(* IEC 61131-3 sources: s7-to-codesys/tests/POUs/Scenarios/FB_Motor_ScenarioTest, 8 files *)

(* ---- FB_Motor_ScenarioTest.decl.st ---- *)
// AUTO-GENERATED — не редактировать: s7conv gen-tests, сценарии scenarios/FB_Motor.csv
// Правка — в CSV (scenarios/README.md), затем python -m s7conv build-corpus.
// Назначение: тесты поведения сконвертированного FB_Motor по сценариям CSV (сценариев: 7, строк: 52):
//             один метод-тест на сценарий, строки — по порядку с моделируемым временем GVL_S7Clock.
//             Ожидаемые значения — из CSV (эталонные модели по описанию логики блока), не из
//             результата конвертации.
// Автор:      s7conv 0.1.0 (сгенерировано)
// Версия:     не указана
// Документ:   scenarios/README.md, docs/methodology.md, раздел «Проверка поведения»
FUNCTION_BLOCK FB_Motor_ScenarioTest EXTENDS coUnit.FB_TestSuite
VAR
    fbAutoStartOk : FB_Motor;  // свой экземпляр на сценарий
    xAutoStartOkDone : BOOL;  // сценарий выполнен (выполняется один раз)
    fbNoFeedbackTimeout : FB_Motor;  // свой экземпляр на сценарий
    xNoFeedbackTimeoutDone : BOOL;  // сценарий выполнен (выполняется один раз)
    fbFeedbackLost : FB_Motor;  // свой экземпляр на сценарий
    xFeedbackLostDone : BOOL;  // сценарий выполнен (выполняется один раз)
    fbUnexpectedFeedback : FB_Motor;  // свой экземпляр на сценарий
    xUnexpectedFeedbackDone : BOOL;  // сценарий выполнен (выполняется один раз)
    fbThermalTripManual : FB_Motor;  // свой экземпляр на сценарий
    xThermalTripManualDone : BOOL;  // сценарий выполнен (выполняется один раз)
    fbBumplessAutoToManual : FB_Motor;  // свой экземпляр на сценарий
    xBumplessAutoToManualDone : BOOL;  // сценарий выполнен (выполняется один раз)
    fbCustomFeedbackTime : FB_Motor;  // свой экземпляр на сценарий
    xCustomFeedbackTimeDone : BOOL;  // сценарий выполнен (выполняется один раз)
END_VAR

(* ---- AutoStartOk.method.impl.st ---- *)
// AUTO-GENERATED — не редактировать: scenarios/FB_Motor.csv, сценарий AutoStartOk
coUnit.TEST('AutoStartOk');
IF NOT xAutoStartOkDone THEN
    xAutoStartOkDone := TRUE;
    GVL_S7Clock.xSimulation := TRUE;

    // #1, t = 0 мс — авто, команды нет
    GVL_S7Clock.tSimNow := T#0MS;
    fbAutoStartOk.autoMode := TRUE;
    fbAutoStartOk.autoStart := FALSE;
    fbAutoStartOk.manStart := FALSE;
    fbAutoStartOk.manStop := FALSE;
    fbAutoStartOk.feedback := FALSE;
    fbAutoStartOk.thermalOk := TRUE;
    fbAutoStartOk.reset := FALSE;
    fbAutoStartOk.feedbackTime := T#3000MS;
    fbAutoStartOk();
    AssertEquals_BOOL(Expected := FALSE, Actual := fbAutoStartOk.runCmd, Message := 'AutoStartOk#1 runCmd');
    AssertEquals_BOOL(Expected := FALSE, Actual := fbAutoStartOk.fault, Message := 'AutoStartOk#1 fault');
    AssertEquals_BOOL(Expected := FALSE,
                      Actual := fbAutoStartOk.status.running,
                      Message := 'AutoStartOk#1 status.running');
    AssertEquals_BOOL(Expected := FALSE, Actual := fbAutoStartOk.status.fault, Message := 'AutoStartOk#1 status.fault');
    AssertEquals_BOOL(Expected := TRUE,
                      Actual := fbAutoStartOk.status.autoMode,
                      Message := 'AutoStartOk#1 status.autoMode');
    AssertEquals_INT(Expected := 0,
                     Actual := fbAutoStartOk.status.faultCode,
                     Message := 'AutoStartOk#1 status.faultCode');
    AssertEquals_DINT(Expected := 0,
                      Actual := fbAutoStartOk.status.startCount,
                      Message := 'AutoStartOk#1 status.startCount');

    // #2, t = 100 мс — пуск: runCmd, пуск №1; таймер рассогласования запущен
    GVL_S7Clock.tSimNow := T#100MS;
    fbAutoStartOk.autoStart := TRUE;
    fbAutoStartOk();
    AssertEquals_BOOL(Expected := TRUE, Actual := fbAutoStartOk.runCmd, Message := 'AutoStartOk#2 runCmd');
    AssertEquals_BOOL(Expected := FALSE, Actual := fbAutoStartOk.fault, Message := 'AutoStartOk#2 fault');
    AssertEquals_BOOL(Expected := FALSE,
                      Actual := fbAutoStartOk.status.running,
                      Message := 'AutoStartOk#2 status.running');
    AssertEquals_BOOL(Expected := FALSE, Actual := fbAutoStartOk.status.fault, Message := 'AutoStartOk#2 status.fault');
    AssertEquals_BOOL(Expected := TRUE,
                      Actual := fbAutoStartOk.status.autoMode,
                      Message := 'AutoStartOk#2 status.autoMode');
    AssertEquals_INT(Expected := 0,
                     Actual := fbAutoStartOk.status.faultCode,
                     Message := 'AutoStartOk#2 status.faultCode');
    AssertEquals_DINT(Expected := 1,
                      Actual := fbAutoStartOk.status.startCount,
                      Message := 'AutoStartOk#2 status.startCount');

    // #3, t = 1100 мс — обратная связь через 1 с: работает
    GVL_S7Clock.tSimNow := T#1100MS;
    fbAutoStartOk.feedback := TRUE;
    fbAutoStartOk();
    AssertEquals_BOOL(Expected := TRUE, Actual := fbAutoStartOk.runCmd, Message := 'AutoStartOk#3 runCmd');
    AssertEquals_BOOL(Expected := FALSE, Actual := fbAutoStartOk.fault, Message := 'AutoStartOk#3 fault');
    AssertEquals_BOOL(Expected := TRUE,
                      Actual := fbAutoStartOk.status.running,
                      Message := 'AutoStartOk#3 status.running');
    AssertEquals_BOOL(Expected := FALSE, Actual := fbAutoStartOk.status.fault, Message := 'AutoStartOk#3 status.fault');
    AssertEquals_BOOL(Expected := TRUE,
                      Actual := fbAutoStartOk.status.autoMode,
                      Message := 'AutoStartOk#3 status.autoMode');
    AssertEquals_INT(Expected := 0,
                     Actual := fbAutoStartOk.status.faultCode,
                     Message := 'AutoStartOk#3 status.faultCode');
    AssertEquals_DINT(Expected := 1,
                      Actual := fbAutoStartOk.status.startCount,
                      Message := 'AutoStartOk#3 status.startCount');

    // #4, t = 5000 мс — работает, аварии нет
    GVL_S7Clock.tSimNow := T#5000MS;
    fbAutoStartOk();
    AssertEquals_BOOL(Expected := TRUE, Actual := fbAutoStartOk.runCmd, Message := 'AutoStartOk#4 runCmd');
    AssertEquals_BOOL(Expected := FALSE, Actual := fbAutoStartOk.fault, Message := 'AutoStartOk#4 fault');
    AssertEquals_BOOL(Expected := TRUE,
                      Actual := fbAutoStartOk.status.running,
                      Message := 'AutoStartOk#4 status.running');
    AssertEquals_BOOL(Expected := FALSE, Actual := fbAutoStartOk.status.fault, Message := 'AutoStartOk#4 status.fault');
    AssertEquals_BOOL(Expected := TRUE,
                      Actual := fbAutoStartOk.status.autoMode,
                      Message := 'AutoStartOk#4 status.autoMode');
    AssertEquals_INT(Expected := 0,
                     Actual := fbAutoStartOk.status.faultCode,
                     Message := 'AutoStartOk#4 status.faultCode');
    AssertEquals_DINT(Expected := 1,
                      Actual := fbAutoStartOk.status.startCount,
                      Message := 'AutoStartOk#4 status.startCount');

    // #5, t = 5100 мс — стоп: runCmd снят, контактор ещё держит — рассогласование
    GVL_S7Clock.tSimNow := T#5100MS;
    fbAutoStartOk.autoStart := FALSE;
    fbAutoStartOk();
    AssertEquals_BOOL(Expected := FALSE, Actual := fbAutoStartOk.runCmd, Message := 'AutoStartOk#5 runCmd');
    AssertEquals_BOOL(Expected := FALSE, Actual := fbAutoStartOk.fault, Message := 'AutoStartOk#5 fault');
    AssertEquals_BOOL(Expected := FALSE,
                      Actual := fbAutoStartOk.status.running,
                      Message := 'AutoStartOk#5 status.running');
    AssertEquals_BOOL(Expected := FALSE, Actual := fbAutoStartOk.status.fault, Message := 'AutoStartOk#5 status.fault');
    AssertEquals_BOOL(Expected := TRUE,
                      Actual := fbAutoStartOk.status.autoMode,
                      Message := 'AutoStartOk#5 status.autoMode');
    AssertEquals_INT(Expected := 0,
                     Actual := fbAutoStartOk.status.faultCode,
                     Message := 'AutoStartOk#5 status.faultCode');
    AssertEquals_DINT(Expected := 1,
                      Actual := fbAutoStartOk.status.startCount,
                      Message := 'AutoStartOk#5 status.startCount');

    // #6, t = 6000 мс — обратная связь пропала через 0.9 с — нормальный останов
    GVL_S7Clock.tSimNow := T#6000MS;
    fbAutoStartOk.feedback := FALSE;
    fbAutoStartOk();
    AssertEquals_BOOL(Expected := FALSE, Actual := fbAutoStartOk.runCmd, Message := 'AutoStartOk#6 runCmd');
    AssertEquals_BOOL(Expected := FALSE, Actual := fbAutoStartOk.fault, Message := 'AutoStartOk#6 fault');
    AssertEquals_BOOL(Expected := FALSE,
                      Actual := fbAutoStartOk.status.running,
                      Message := 'AutoStartOk#6 status.running');
    AssertEquals_BOOL(Expected := FALSE, Actual := fbAutoStartOk.status.fault, Message := 'AutoStartOk#6 status.fault');
    AssertEquals_BOOL(Expected := TRUE,
                      Actual := fbAutoStartOk.status.autoMode,
                      Message := 'AutoStartOk#6 status.autoMode');
    AssertEquals_INT(Expected := 0,
                     Actual := fbAutoStartOk.status.faultCode,
                     Message := 'AutoStartOk#6 status.faultCode');
    AssertEquals_DINT(Expected := 1,
                      Actual := fbAutoStartOk.status.startCount,
                      Message := 'AutoStartOk#6 status.startCount');

    // #7, t = 9500 мс — покой
    GVL_S7Clock.tSimNow := T#9500MS;
    fbAutoStartOk();
    AssertEquals_BOOL(Expected := FALSE, Actual := fbAutoStartOk.runCmd, Message := 'AutoStartOk#7 runCmd');
    AssertEquals_BOOL(Expected := FALSE, Actual := fbAutoStartOk.fault, Message := 'AutoStartOk#7 fault');
    AssertEquals_BOOL(Expected := FALSE,
                      Actual := fbAutoStartOk.status.running,
                      Message := 'AutoStartOk#7 status.running');
    AssertEquals_BOOL(Expected := FALSE, Actual := fbAutoStartOk.status.fault, Message := 'AutoStartOk#7 status.fault');
    AssertEquals_BOOL(Expected := TRUE,
                      Actual := fbAutoStartOk.status.autoMode,
                      Message := 'AutoStartOk#7 status.autoMode');
    AssertEquals_INT(Expected := 0,
                     Actual := fbAutoStartOk.status.faultCode,
                     Message := 'AutoStartOk#7 status.faultCode');
    AssertEquals_DINT(Expected := 1,
                      Actual := fbAutoStartOk.status.startCount,
                      Message := 'AutoStartOk#7 status.startCount');

    GVL_S7Clock.xSimulation := FALSE;
END_IF
coUnit.TEST_FINISHED();

(* ---- BumplessAutoToManual.method.impl.st ---- *)
// AUTO-GENERATED — не редактировать: scenarios/FB_Motor.csv, сценарий BumplessAutoToManual
coUnit.TEST('BumplessAutoToManual');
IF NOT xBumplessAutoToManualDone THEN
    xBumplessAutoToManualDone := TRUE;
    GVL_S7Clock.xSimulation := TRUE;

    // #1, t = 0 мс — авто, пуск №1
    GVL_S7Clock.tSimNow := T#0MS;
    fbBumplessAutoToManual.autoMode := TRUE;
    fbBumplessAutoToManual.autoStart := TRUE;
    fbBumplessAutoToManual.manStart := FALSE;
    fbBumplessAutoToManual.manStop := FALSE;
    fbBumplessAutoToManual.feedback := FALSE;
    fbBumplessAutoToManual.thermalOk := TRUE;
    fbBumplessAutoToManual.reset := FALSE;
    fbBumplessAutoToManual.feedbackTime := T#3000MS;
    fbBumplessAutoToManual();
    AssertEquals_BOOL(Expected := TRUE,
                      Actual := fbBumplessAutoToManual.runCmd,
                      Message := 'BumplessAutoToManual#1 runCmd');
    AssertEquals_BOOL(Expected := FALSE,
                      Actual := fbBumplessAutoToManual.fault,
                      Message := 'BumplessAutoToManual#1 fault');
    AssertEquals_BOOL(Expected := FALSE,
                      Actual := fbBumplessAutoToManual.status.running,
                      Message := 'BumplessAutoToManual#1 status.running');
    AssertEquals_BOOL(Expected := FALSE,
                      Actual := fbBumplessAutoToManual.status.fault,
                      Message := 'BumplessAutoToManual#1 status.fault');
    AssertEquals_BOOL(Expected := TRUE,
                      Actual := fbBumplessAutoToManual.status.autoMode,
                      Message := 'BumplessAutoToManual#1 status.autoMode');
    AssertEquals_INT(Expected := 0,
                     Actual := fbBumplessAutoToManual.status.faultCode,
                     Message := 'BumplessAutoToManual#1 status.faultCode');
    AssertEquals_DINT(Expected := 1,
                      Actual := fbBumplessAutoToManual.status.startCount,
                      Message := 'BumplessAutoToManual#1 status.startCount');

    // #2, t = 500 мс — работает
    GVL_S7Clock.tSimNow := T#500MS;
    fbBumplessAutoToManual.feedback := TRUE;
    fbBumplessAutoToManual();
    AssertEquals_BOOL(Expected := TRUE,
                      Actual := fbBumplessAutoToManual.runCmd,
                      Message := 'BumplessAutoToManual#2 runCmd');
    AssertEquals_BOOL(Expected := FALSE,
                      Actual := fbBumplessAutoToManual.fault,
                      Message := 'BumplessAutoToManual#2 fault');
    AssertEquals_BOOL(Expected := TRUE,
                      Actual := fbBumplessAutoToManual.status.running,
                      Message := 'BumplessAutoToManual#2 status.running');
    AssertEquals_BOOL(Expected := FALSE,
                      Actual := fbBumplessAutoToManual.status.fault,
                      Message := 'BumplessAutoToManual#2 status.fault');
    AssertEquals_BOOL(Expected := TRUE,
                      Actual := fbBumplessAutoToManual.status.autoMode,
                      Message := 'BumplessAutoToManual#2 status.autoMode');
    AssertEquals_INT(Expected := 0,
                     Actual := fbBumplessAutoToManual.status.faultCode,
                     Message := 'BumplessAutoToManual#2 status.faultCode');
    AssertEquals_DINT(Expected := 1,
                      Actual := fbBumplessAutoToManual.status.startCount,
                      Message := 'BumplessAutoToManual#2 status.startCount');

    // #3, t = 1000 мс — в ручной: защёлка следила за авто — продолжает работать
    GVL_S7Clock.tSimNow := T#1000MS;
    fbBumplessAutoToManual.autoMode := FALSE;
    fbBumplessAutoToManual();
    AssertEquals_BOOL(Expected := TRUE,
                      Actual := fbBumplessAutoToManual.runCmd,
                      Message := 'BumplessAutoToManual#3 runCmd');
    AssertEquals_BOOL(Expected := FALSE,
                      Actual := fbBumplessAutoToManual.fault,
                      Message := 'BumplessAutoToManual#3 fault');
    AssertEquals_BOOL(Expected := TRUE,
                      Actual := fbBumplessAutoToManual.status.running,
                      Message := 'BumplessAutoToManual#3 status.running');
    AssertEquals_BOOL(Expected := FALSE,
                      Actual := fbBumplessAutoToManual.status.fault,
                      Message := 'BumplessAutoToManual#3 status.fault');
    AssertEquals_BOOL(Expected := FALSE,
                      Actual := fbBumplessAutoToManual.status.autoMode,
                      Message := 'BumplessAutoToManual#3 status.autoMode');
    AssertEquals_INT(Expected := 0,
                     Actual := fbBumplessAutoToManual.status.faultCode,
                     Message := 'BumplessAutoToManual#3 status.faultCode');
    AssertEquals_DINT(Expected := 1,
                      Actual := fbBumplessAutoToManual.status.startCount,
                      Message := 'BumplessAutoToManual#3 status.startCount');

    // #4, t = 2000 мс — стоп оператором
    GVL_S7Clock.tSimNow := T#2000MS;
    fbBumplessAutoToManual.manStop := TRUE;
    fbBumplessAutoToManual();
    AssertEquals_BOOL(Expected := FALSE,
                      Actual := fbBumplessAutoToManual.runCmd,
                      Message := 'BumplessAutoToManual#4 runCmd');
    AssertEquals_BOOL(Expected := FALSE,
                      Actual := fbBumplessAutoToManual.fault,
                      Message := 'BumplessAutoToManual#4 fault');
    AssertEquals_BOOL(Expected := FALSE,
                      Actual := fbBumplessAutoToManual.status.running,
                      Message := 'BumplessAutoToManual#4 status.running');
    AssertEquals_BOOL(Expected := FALSE,
                      Actual := fbBumplessAutoToManual.status.fault,
                      Message := 'BumplessAutoToManual#4 status.fault');
    AssertEquals_BOOL(Expected := FALSE,
                      Actual := fbBumplessAutoToManual.status.autoMode,
                      Message := 'BumplessAutoToManual#4 status.autoMode');
    AssertEquals_INT(Expected := 0,
                     Actual := fbBumplessAutoToManual.status.faultCode,
                     Message := 'BumplessAutoToManual#4 status.faultCode');
    AssertEquals_DINT(Expected := 1,
                      Actual := fbBumplessAutoToManual.status.startCount,
                      Message := 'BumplessAutoToManual#4 status.startCount');

    // #5, t = 2500 мс — остановлен
    GVL_S7Clock.tSimNow := T#2500MS;
    fbBumplessAutoToManual.manStop := FALSE;
    fbBumplessAutoToManual.feedback := FALSE;
    fbBumplessAutoToManual();
    AssertEquals_BOOL(Expected := FALSE,
                      Actual := fbBumplessAutoToManual.runCmd,
                      Message := 'BumplessAutoToManual#5 runCmd');
    AssertEquals_BOOL(Expected := FALSE,
                      Actual := fbBumplessAutoToManual.fault,
                      Message := 'BumplessAutoToManual#5 fault');
    AssertEquals_BOOL(Expected := FALSE,
                      Actual := fbBumplessAutoToManual.status.running,
                      Message := 'BumplessAutoToManual#5 status.running');
    AssertEquals_BOOL(Expected := FALSE,
                      Actual := fbBumplessAutoToManual.status.fault,
                      Message := 'BumplessAutoToManual#5 status.fault');
    AssertEquals_BOOL(Expected := FALSE,
                      Actual := fbBumplessAutoToManual.status.autoMode,
                      Message := 'BumplessAutoToManual#5 status.autoMode');
    AssertEquals_INT(Expected := 0,
                     Actual := fbBumplessAutoToManual.status.faultCode,
                     Message := 'BumplessAutoToManual#5 status.faultCode');
    AssertEquals_DINT(Expected := 1,
                      Actual := fbBumplessAutoToManual.status.startCount,
                      Message := 'BumplessAutoToManual#5 status.startCount');

    // #6, t = 3000 мс — в авто без запроса
    GVL_S7Clock.tSimNow := T#3000MS;
    fbBumplessAutoToManual.autoMode := TRUE;
    fbBumplessAutoToManual.autoStart := FALSE;
    fbBumplessAutoToManual();
    AssertEquals_BOOL(Expected := FALSE,
                      Actual := fbBumplessAutoToManual.runCmd,
                      Message := 'BumplessAutoToManual#6 runCmd');
    AssertEquals_BOOL(Expected := FALSE,
                      Actual := fbBumplessAutoToManual.fault,
                      Message := 'BumplessAutoToManual#6 fault');
    AssertEquals_BOOL(Expected := FALSE,
                      Actual := fbBumplessAutoToManual.status.running,
                      Message := 'BumplessAutoToManual#6 status.running');
    AssertEquals_BOOL(Expected := FALSE,
                      Actual := fbBumplessAutoToManual.status.fault,
                      Message := 'BumplessAutoToManual#6 status.fault');
    AssertEquals_BOOL(Expected := TRUE,
                      Actual := fbBumplessAutoToManual.status.autoMode,
                      Message := 'BumplessAutoToManual#6 status.autoMode');
    AssertEquals_INT(Expected := 0,
                     Actual := fbBumplessAutoToManual.status.faultCode,
                     Message := 'BumplessAutoToManual#6 status.faultCode');
    AssertEquals_DINT(Expected := 1,
                      Actual := fbBumplessAutoToManual.status.startCount,
                      Message := 'BumplessAutoToManual#6 status.startCount');

    // #7, t = 3500 мс — запрос авто: пуск №2
    GVL_S7Clock.tSimNow := T#3500MS;
    fbBumplessAutoToManual.autoStart := TRUE;
    fbBumplessAutoToManual();
    AssertEquals_BOOL(Expected := TRUE,
                      Actual := fbBumplessAutoToManual.runCmd,
                      Message := 'BumplessAutoToManual#7 runCmd');
    AssertEquals_BOOL(Expected := FALSE,
                      Actual := fbBumplessAutoToManual.fault,
                      Message := 'BumplessAutoToManual#7 fault');
    AssertEquals_BOOL(Expected := FALSE,
                      Actual := fbBumplessAutoToManual.status.running,
                      Message := 'BumplessAutoToManual#7 status.running');
    AssertEquals_BOOL(Expected := FALSE,
                      Actual := fbBumplessAutoToManual.status.fault,
                      Message := 'BumplessAutoToManual#7 status.fault');
    AssertEquals_BOOL(Expected := TRUE,
                      Actual := fbBumplessAutoToManual.status.autoMode,
                      Message := 'BumplessAutoToManual#7 status.autoMode');
    AssertEquals_INT(Expected := 0,
                     Actual := fbBumplessAutoToManual.status.faultCode,
                     Message := 'BumplessAutoToManual#7 status.faultCode');
    AssertEquals_DINT(Expected := 2,
                      Actual := fbBumplessAutoToManual.status.startCount,
                      Message := 'BumplessAutoToManual#7 status.startCount');

    // #8, t = 4000 мс — работает
    GVL_S7Clock.tSimNow := T#4000MS;
    fbBumplessAutoToManual.feedback := TRUE;
    fbBumplessAutoToManual();
    AssertEquals_BOOL(Expected := TRUE,
                      Actual := fbBumplessAutoToManual.runCmd,
                      Message := 'BumplessAutoToManual#8 runCmd');
    AssertEquals_BOOL(Expected := FALSE,
                      Actual := fbBumplessAutoToManual.fault,
                      Message := 'BumplessAutoToManual#8 fault');
    AssertEquals_BOOL(Expected := TRUE,
                      Actual := fbBumplessAutoToManual.status.running,
                      Message := 'BumplessAutoToManual#8 status.running');
    AssertEquals_BOOL(Expected := FALSE,
                      Actual := fbBumplessAutoToManual.status.fault,
                      Message := 'BumplessAutoToManual#8 status.fault');
    AssertEquals_BOOL(Expected := TRUE,
                      Actual := fbBumplessAutoToManual.status.autoMode,
                      Message := 'BumplessAutoToManual#8 status.autoMode');
    AssertEquals_INT(Expected := 0,
                     Actual := fbBumplessAutoToManual.status.faultCode,
                     Message := 'BumplessAutoToManual#8 status.faultCode');
    AssertEquals_DINT(Expected := 2,
                      Actual := fbBumplessAutoToManual.status.startCount,
                      Message := 'BumplessAutoToManual#8 status.startCount');

    GVL_S7Clock.xSimulation := FALSE;
END_IF
coUnit.TEST_FINISHED();

(* ---- CustomFeedbackTime.method.impl.st ---- *)
// AUTO-GENERATED — не редактировать: scenarios/FB_Motor.csv, сценарий CustomFeedbackTime
coUnit.TEST('CustomFeedbackTime');
IF NOT xCustomFeedbackTimeDone THEN
    xCustomFeedbackTimeDone := TRUE;
    GVL_S7Clock.xSimulation := TRUE;

    // #1, t = 0 мс — пуск, feedbackTime 5 с
    GVL_S7Clock.tSimNow := T#0MS;
    fbCustomFeedbackTime.autoMode := TRUE;
    fbCustomFeedbackTime.autoStart := TRUE;
    fbCustomFeedbackTime.manStart := FALSE;
    fbCustomFeedbackTime.manStop := FALSE;
    fbCustomFeedbackTime.feedback := FALSE;
    fbCustomFeedbackTime.thermalOk := TRUE;
    fbCustomFeedbackTime.reset := FALSE;
    fbCustomFeedbackTime.feedbackTime := T#5000MS;
    fbCustomFeedbackTime();
    AssertEquals_BOOL(Expected := TRUE,
                      Actual := fbCustomFeedbackTime.runCmd,
                      Message := 'CustomFeedbackTime#1 runCmd');
    AssertEquals_BOOL(Expected := FALSE, Actual := fbCustomFeedbackTime.fault, Message := 'CustomFeedbackTime#1 fault');
    AssertEquals_BOOL(Expected := FALSE,
                      Actual := fbCustomFeedbackTime.status.running,
                      Message := 'CustomFeedbackTime#1 status.running');
    AssertEquals_BOOL(Expected := FALSE,
                      Actual := fbCustomFeedbackTime.status.fault,
                      Message := 'CustomFeedbackTime#1 status.fault');
    AssertEquals_BOOL(Expected := TRUE,
                      Actual := fbCustomFeedbackTime.status.autoMode,
                      Message := 'CustomFeedbackTime#1 status.autoMode');
    AssertEquals_INT(Expected := 0,
                     Actual := fbCustomFeedbackTime.status.faultCode,
                     Message := 'CustomFeedbackTime#1 status.faultCode');
    AssertEquals_DINT(Expected := 1,
                      Actual := fbCustomFeedbackTime.status.startCount,
                      Message := 'CustomFeedbackTime#1 status.startCount');

    // #2, t = 4500 мс — обратная связь через 4.5 с — аварии нет
    GVL_S7Clock.tSimNow := T#4500MS;
    fbCustomFeedbackTime.feedback := TRUE;
    fbCustomFeedbackTime();
    AssertEquals_BOOL(Expected := TRUE,
                      Actual := fbCustomFeedbackTime.runCmd,
                      Message := 'CustomFeedbackTime#2 runCmd');
    AssertEquals_BOOL(Expected := FALSE, Actual := fbCustomFeedbackTime.fault, Message := 'CustomFeedbackTime#2 fault');
    AssertEquals_BOOL(Expected := TRUE,
                      Actual := fbCustomFeedbackTime.status.running,
                      Message := 'CustomFeedbackTime#2 status.running');
    AssertEquals_BOOL(Expected := FALSE,
                      Actual := fbCustomFeedbackTime.status.fault,
                      Message := 'CustomFeedbackTime#2 status.fault');
    AssertEquals_BOOL(Expected := TRUE,
                      Actual := fbCustomFeedbackTime.status.autoMode,
                      Message := 'CustomFeedbackTime#2 status.autoMode');
    AssertEquals_INT(Expected := 0,
                     Actual := fbCustomFeedbackTime.status.faultCode,
                     Message := 'CustomFeedbackTime#2 status.faultCode');
    AssertEquals_DINT(Expected := 1,
                      Actual := fbCustomFeedbackTime.status.startCount,
                      Message := 'CustomFeedbackTime#2 status.startCount');

    // #3, t = 6000 мс — работает
    GVL_S7Clock.tSimNow := T#6000MS;
    fbCustomFeedbackTime();
    AssertEquals_BOOL(Expected := TRUE,
                      Actual := fbCustomFeedbackTime.runCmd,
                      Message := 'CustomFeedbackTime#3 runCmd');
    AssertEquals_BOOL(Expected := FALSE, Actual := fbCustomFeedbackTime.fault, Message := 'CustomFeedbackTime#3 fault');
    AssertEquals_BOOL(Expected := TRUE,
                      Actual := fbCustomFeedbackTime.status.running,
                      Message := 'CustomFeedbackTime#3 status.running');
    AssertEquals_BOOL(Expected := FALSE,
                      Actual := fbCustomFeedbackTime.status.fault,
                      Message := 'CustomFeedbackTime#3 status.fault');
    AssertEquals_BOOL(Expected := TRUE,
                      Actual := fbCustomFeedbackTime.status.autoMode,
                      Message := 'CustomFeedbackTime#3 status.autoMode');
    AssertEquals_INT(Expected := 0,
                     Actual := fbCustomFeedbackTime.status.faultCode,
                     Message := 'CustomFeedbackTime#3 status.faultCode');
    AssertEquals_DINT(Expected := 1,
                      Actual := fbCustomFeedbackTime.status.startCount,
                      Message := 'CustomFeedbackTime#3 status.startCount');

    GVL_S7Clock.xSimulation := FALSE;
END_IF
coUnit.TEST_FINISHED();

(* ---- FeedbackLost.method.impl.st ---- *)
// AUTO-GENERATED — не редактировать: scenarios/FB_Motor.csv, сценарий FeedbackLost
coUnit.TEST('FeedbackLost');
IF NOT xFeedbackLostDone THEN
    xFeedbackLostDone := TRUE;
    GVL_S7Clock.xSimulation := TRUE;

    // #1, t = 0 мс — пуск
    GVL_S7Clock.tSimNow := T#0MS;
    fbFeedbackLost.autoMode := TRUE;
    fbFeedbackLost.autoStart := TRUE;
    fbFeedbackLost.manStart := FALSE;
    fbFeedbackLost.manStop := FALSE;
    fbFeedbackLost.feedback := FALSE;
    fbFeedbackLost.thermalOk := TRUE;
    fbFeedbackLost.reset := FALSE;
    fbFeedbackLost.feedbackTime := T#3000MS;
    fbFeedbackLost();
    AssertEquals_BOOL(Expected := TRUE, Actual := fbFeedbackLost.runCmd, Message := 'FeedbackLost#1 runCmd');
    AssertEquals_BOOL(Expected := FALSE, Actual := fbFeedbackLost.fault, Message := 'FeedbackLost#1 fault');
    AssertEquals_BOOL(Expected := FALSE,
                      Actual := fbFeedbackLost.status.running,
                      Message := 'FeedbackLost#1 status.running');
    AssertEquals_BOOL(Expected := FALSE,
                      Actual := fbFeedbackLost.status.fault,
                      Message := 'FeedbackLost#1 status.fault');
    AssertEquals_BOOL(Expected := TRUE,
                      Actual := fbFeedbackLost.status.autoMode,
                      Message := 'FeedbackLost#1 status.autoMode');
    AssertEquals_INT(Expected := 0,
                     Actual := fbFeedbackLost.status.faultCode,
                     Message := 'FeedbackLost#1 status.faultCode');
    AssertEquals_DINT(Expected := 1,
                      Actual := fbFeedbackLost.status.startCount,
                      Message := 'FeedbackLost#1 status.startCount');

    // #2, t = 500 мс — обратная связь есть
    GVL_S7Clock.tSimNow := T#500MS;
    fbFeedbackLost.feedback := TRUE;
    fbFeedbackLost();
    AssertEquals_BOOL(Expected := TRUE, Actual := fbFeedbackLost.runCmd, Message := 'FeedbackLost#2 runCmd');
    AssertEquals_BOOL(Expected := FALSE, Actual := fbFeedbackLost.fault, Message := 'FeedbackLost#2 fault');
    AssertEquals_BOOL(Expected := TRUE,
                      Actual := fbFeedbackLost.status.running,
                      Message := 'FeedbackLost#2 status.running');
    AssertEquals_BOOL(Expected := FALSE,
                      Actual := fbFeedbackLost.status.fault,
                      Message := 'FeedbackLost#2 status.fault');
    AssertEquals_BOOL(Expected := TRUE,
                      Actual := fbFeedbackLost.status.autoMode,
                      Message := 'FeedbackLost#2 status.autoMode');
    AssertEquals_INT(Expected := 0,
                     Actual := fbFeedbackLost.status.faultCode,
                     Message := 'FeedbackLost#2 status.faultCode');
    AssertEquals_DINT(Expected := 1,
                      Actual := fbFeedbackLost.status.startCount,
                      Message := 'FeedbackLost#2 status.startCount');

    // #3, t = 10000 мс — обратная связь пропала; отсчёт с 10.0 с
    GVL_S7Clock.tSimNow := T#10000MS;
    fbFeedbackLost.feedback := FALSE;
    fbFeedbackLost();
    AssertEquals_BOOL(Expected := TRUE, Actual := fbFeedbackLost.runCmd, Message := 'FeedbackLost#3 runCmd');
    AssertEquals_BOOL(Expected := FALSE, Actual := fbFeedbackLost.fault, Message := 'FeedbackLost#3 fault');
    AssertEquals_BOOL(Expected := FALSE,
                      Actual := fbFeedbackLost.status.running,
                      Message := 'FeedbackLost#3 status.running');
    AssertEquals_BOOL(Expected := FALSE,
                      Actual := fbFeedbackLost.status.fault,
                      Message := 'FeedbackLost#3 status.fault');
    AssertEquals_BOOL(Expected := TRUE,
                      Actual := fbFeedbackLost.status.autoMode,
                      Message := 'FeedbackLost#3 status.autoMode');
    AssertEquals_INT(Expected := 0,
                     Actual := fbFeedbackLost.status.faultCode,
                     Message := 'FeedbackLost#3 status.faultCode');
    AssertEquals_DINT(Expected := 1,
                      Actual := fbFeedbackLost.status.startCount,
                      Message := 'FeedbackLost#3 status.startCount');

    // #4, t = 12800 мс — 2.8 с без обратной связи: аварии нет
    GVL_S7Clock.tSimNow := T#12800MS;
    fbFeedbackLost();
    AssertEquals_BOOL(Expected := TRUE, Actual := fbFeedbackLost.runCmd, Message := 'FeedbackLost#4 runCmd');
    AssertEquals_BOOL(Expected := FALSE, Actual := fbFeedbackLost.fault, Message := 'FeedbackLost#4 fault');
    AssertEquals_BOOL(Expected := FALSE,
                      Actual := fbFeedbackLost.status.running,
                      Message := 'FeedbackLost#4 status.running');
    AssertEquals_BOOL(Expected := FALSE,
                      Actual := fbFeedbackLost.status.fault,
                      Message := 'FeedbackLost#4 status.fault');
    AssertEquals_BOOL(Expected := TRUE,
                      Actual := fbFeedbackLost.status.autoMode,
                      Message := 'FeedbackLost#4 status.autoMode');
    AssertEquals_INT(Expected := 0,
                     Actual := fbFeedbackLost.status.faultCode,
                     Message := 'FeedbackLost#4 status.faultCode');
    AssertEquals_DINT(Expected := 1,
                      Actual := fbFeedbackLost.status.startCount,
                      Message := 'FeedbackLost#4 status.startCount');

    // #5, t = 13200 мс — 3.2 с: авария 2 (обратная связь уже была), runCmd снят
    GVL_S7Clock.tSimNow := T#13200MS;
    fbFeedbackLost();
    AssertEquals_BOOL(Expected := FALSE, Actual := fbFeedbackLost.runCmd, Message := 'FeedbackLost#5 runCmd');
    AssertEquals_BOOL(Expected := TRUE, Actual := fbFeedbackLost.fault, Message := 'FeedbackLost#5 fault');
    AssertEquals_BOOL(Expected := FALSE,
                      Actual := fbFeedbackLost.status.running,
                      Message := 'FeedbackLost#5 status.running');
    AssertEquals_BOOL(Expected := TRUE,
                      Actual := fbFeedbackLost.status.fault,
                      Message := 'FeedbackLost#5 status.fault');
    AssertEquals_BOOL(Expected := TRUE,
                      Actual := fbFeedbackLost.status.autoMode,
                      Message := 'FeedbackLost#5 status.autoMode');
    AssertEquals_INT(Expected := 2,
                     Actual := fbFeedbackLost.status.faultCode,
                     Message := 'FeedbackLost#5 status.faultCode');
    AssertEquals_DINT(Expected := 1,
                      Actual := fbFeedbackLost.status.startCount,
                      Message := 'FeedbackLost#5 status.startCount');

    // #6, t = 14000 мс — сброс, запроса нет — стоит без аварии
    GVL_S7Clock.tSimNow := T#14000MS;
    fbFeedbackLost.autoStart := FALSE;
    fbFeedbackLost.reset := TRUE;
    fbFeedbackLost();
    AssertEquals_BOOL(Expected := FALSE, Actual := fbFeedbackLost.runCmd, Message := 'FeedbackLost#6 runCmd');
    AssertEquals_BOOL(Expected := FALSE, Actual := fbFeedbackLost.fault, Message := 'FeedbackLost#6 fault');
    AssertEquals_BOOL(Expected := FALSE,
                      Actual := fbFeedbackLost.status.running,
                      Message := 'FeedbackLost#6 status.running');
    AssertEquals_BOOL(Expected := FALSE,
                      Actual := fbFeedbackLost.status.fault,
                      Message := 'FeedbackLost#6 status.fault');
    AssertEquals_BOOL(Expected := TRUE,
                      Actual := fbFeedbackLost.status.autoMode,
                      Message := 'FeedbackLost#6 status.autoMode');
    AssertEquals_INT(Expected := 0,
                     Actual := fbFeedbackLost.status.faultCode,
                     Message := 'FeedbackLost#6 status.faultCode');
    AssertEquals_DINT(Expected := 1,
                      Actual := fbFeedbackLost.status.startCount,
                      Message := 'FeedbackLost#6 status.startCount');

    // #7, t = 14500 мс — покой
    GVL_S7Clock.tSimNow := T#14500MS;
    fbFeedbackLost.reset := FALSE;
    fbFeedbackLost();
    AssertEquals_BOOL(Expected := FALSE, Actual := fbFeedbackLost.runCmd, Message := 'FeedbackLost#7 runCmd');
    AssertEquals_BOOL(Expected := FALSE, Actual := fbFeedbackLost.fault, Message := 'FeedbackLost#7 fault');
    AssertEquals_BOOL(Expected := FALSE,
                      Actual := fbFeedbackLost.status.running,
                      Message := 'FeedbackLost#7 status.running');
    AssertEquals_BOOL(Expected := FALSE,
                      Actual := fbFeedbackLost.status.fault,
                      Message := 'FeedbackLost#7 status.fault');
    AssertEquals_BOOL(Expected := TRUE,
                      Actual := fbFeedbackLost.status.autoMode,
                      Message := 'FeedbackLost#7 status.autoMode');
    AssertEquals_INT(Expected := 0,
                     Actual := fbFeedbackLost.status.faultCode,
                     Message := 'FeedbackLost#7 status.faultCode');
    AssertEquals_DINT(Expected := 1,
                      Actual := fbFeedbackLost.status.startCount,
                      Message := 'FeedbackLost#7 status.startCount');

    GVL_S7Clock.xSimulation := FALSE;
END_IF
coUnit.TEST_FINISHED();

(* ---- NoFeedbackTimeout.method.impl.st ---- *)
// AUTO-GENERATED — не редактировать: scenarios/FB_Motor.csv, сценарий NoFeedbackTimeout
coUnit.TEST('NoFeedbackTimeout');
IF NOT xNoFeedbackTimeoutDone THEN
    xNoFeedbackTimeoutDone := TRUE;
    GVL_S7Clock.xSimulation := TRUE;

    // #1, t = 0 мс — пуск, обратной связи нет
    GVL_S7Clock.tSimNow := T#0MS;
    fbNoFeedbackTimeout.autoMode := TRUE;
    fbNoFeedbackTimeout.autoStart := TRUE;
    fbNoFeedbackTimeout.manStart := FALSE;
    fbNoFeedbackTimeout.manStop := FALSE;
    fbNoFeedbackTimeout.feedback := FALSE;
    fbNoFeedbackTimeout.thermalOk := TRUE;
    fbNoFeedbackTimeout.reset := FALSE;
    fbNoFeedbackTimeout.feedbackTime := T#3000MS;
    fbNoFeedbackTimeout();
    AssertEquals_BOOL(Expected := TRUE, Actual := fbNoFeedbackTimeout.runCmd, Message := 'NoFeedbackTimeout#1 runCmd');
    AssertEquals_BOOL(Expected := FALSE, Actual := fbNoFeedbackTimeout.fault, Message := 'NoFeedbackTimeout#1 fault');
    AssertEquals_BOOL(Expected := FALSE,
                      Actual := fbNoFeedbackTimeout.status.running,
                      Message := 'NoFeedbackTimeout#1 status.running');
    AssertEquals_BOOL(Expected := FALSE,
                      Actual := fbNoFeedbackTimeout.status.fault,
                      Message := 'NoFeedbackTimeout#1 status.fault');
    AssertEquals_BOOL(Expected := TRUE,
                      Actual := fbNoFeedbackTimeout.status.autoMode,
                      Message := 'NoFeedbackTimeout#1 status.autoMode');
    AssertEquals_INT(Expected := 0,
                     Actual := fbNoFeedbackTimeout.status.faultCode,
                     Message := 'NoFeedbackTimeout#1 status.faultCode');
    AssertEquals_DINT(Expected := 1,
                      Actual := fbNoFeedbackTimeout.status.startCount,
                      Message := 'NoFeedbackTimeout#1 status.startCount');

    // #2, t = 2800 мс — 2.8 с < 3 с: аварии нет
    GVL_S7Clock.tSimNow := T#2800MS;
    fbNoFeedbackTimeout();
    AssertEquals_BOOL(Expected := TRUE, Actual := fbNoFeedbackTimeout.runCmd, Message := 'NoFeedbackTimeout#2 runCmd');
    AssertEquals_BOOL(Expected := FALSE, Actual := fbNoFeedbackTimeout.fault, Message := 'NoFeedbackTimeout#2 fault');
    AssertEquals_BOOL(Expected := FALSE,
                      Actual := fbNoFeedbackTimeout.status.running,
                      Message := 'NoFeedbackTimeout#2 status.running');
    AssertEquals_BOOL(Expected := FALSE,
                      Actual := fbNoFeedbackTimeout.status.fault,
                      Message := 'NoFeedbackTimeout#2 status.fault');
    AssertEquals_BOOL(Expected := TRUE,
                      Actual := fbNoFeedbackTimeout.status.autoMode,
                      Message := 'NoFeedbackTimeout#2 status.autoMode');
    AssertEquals_INT(Expected := 0,
                     Actual := fbNoFeedbackTimeout.status.faultCode,
                     Message := 'NoFeedbackTimeout#2 status.faultCode');
    AssertEquals_DINT(Expected := 1,
                      Actual := fbNoFeedbackTimeout.status.startCount,
                      Message := 'NoFeedbackTimeout#2 status.startCount');

    // #3, t = 3000 мс, на пороге таймера — 3.0 с = feedbackTime: авария 1, runCmd снят в этом же вызове
    GVL_S7Clock.tSimNow := T#3000MS;
    fbNoFeedbackTimeout();
    AssertEquals_BOOL(Expected := FALSE, Actual := fbNoFeedbackTimeout.runCmd, Message := 'NoFeedbackTimeout#3 runCmd');
    AssertEquals_BOOL(Expected := TRUE, Actual := fbNoFeedbackTimeout.fault, Message := 'NoFeedbackTimeout#3 fault');
    AssertEquals_BOOL(Expected := FALSE,
                      Actual := fbNoFeedbackTimeout.status.running,
                      Message := 'NoFeedbackTimeout#3 status.running');
    AssertEquals_BOOL(Expected := TRUE,
                      Actual := fbNoFeedbackTimeout.status.fault,
                      Message := 'NoFeedbackTimeout#3 status.fault');
    AssertEquals_BOOL(Expected := TRUE,
                      Actual := fbNoFeedbackTimeout.status.autoMode,
                      Message := 'NoFeedbackTimeout#3 status.autoMode');
    AssertEquals_INT(Expected := 1,
                     Actual := fbNoFeedbackTimeout.status.faultCode,
                     Message := 'NoFeedbackTimeout#3 status.faultCode');
    AssertEquals_DINT(Expected := 1,
                      Actual := fbNoFeedbackTimeout.status.startCount,
                      Message := 'NoFeedbackTimeout#3 status.startCount');

    // #4, t = 3200 мс — авария держится, код 1
    GVL_S7Clock.tSimNow := T#3200MS;
    fbNoFeedbackTimeout();
    AssertEquals_BOOL(Expected := FALSE, Actual := fbNoFeedbackTimeout.runCmd, Message := 'NoFeedbackTimeout#4 runCmd');
    AssertEquals_BOOL(Expected := TRUE, Actual := fbNoFeedbackTimeout.fault, Message := 'NoFeedbackTimeout#4 fault');
    AssertEquals_BOOL(Expected := FALSE,
                      Actual := fbNoFeedbackTimeout.status.running,
                      Message := 'NoFeedbackTimeout#4 status.running');
    AssertEquals_BOOL(Expected := TRUE,
                      Actual := fbNoFeedbackTimeout.status.fault,
                      Message := 'NoFeedbackTimeout#4 status.fault');
    AssertEquals_BOOL(Expected := TRUE,
                      Actual := fbNoFeedbackTimeout.status.autoMode,
                      Message := 'NoFeedbackTimeout#4 status.autoMode');
    AssertEquals_INT(Expected := 1,
                     Actual := fbNoFeedbackTimeout.status.faultCode,
                     Message := 'NoFeedbackTimeout#4 status.faultCode');
    AssertEquals_DINT(Expected := 1,
                      Actual := fbNoFeedbackTimeout.status.startCount,
                      Message := 'NoFeedbackTimeout#4 status.startCount');

    // #5, t = 4000 мс — сброс по фронту: авто-запрос ещё есть — повторный пуск №2
    GVL_S7Clock.tSimNow := T#4000MS;
    fbNoFeedbackTimeout.reset := TRUE;
    fbNoFeedbackTimeout();
    AssertEquals_BOOL(Expected := TRUE, Actual := fbNoFeedbackTimeout.runCmd, Message := 'NoFeedbackTimeout#5 runCmd');
    AssertEquals_BOOL(Expected := FALSE, Actual := fbNoFeedbackTimeout.fault, Message := 'NoFeedbackTimeout#5 fault');
    AssertEquals_BOOL(Expected := FALSE,
                      Actual := fbNoFeedbackTimeout.status.running,
                      Message := 'NoFeedbackTimeout#5 status.running');
    AssertEquals_BOOL(Expected := FALSE,
                      Actual := fbNoFeedbackTimeout.status.fault,
                      Message := 'NoFeedbackTimeout#5 status.fault');
    AssertEquals_BOOL(Expected := TRUE,
                      Actual := fbNoFeedbackTimeout.status.autoMode,
                      Message := 'NoFeedbackTimeout#5 status.autoMode');
    AssertEquals_INT(Expected := 0,
                     Actual := fbNoFeedbackTimeout.status.faultCode,
                     Message := 'NoFeedbackTimeout#5 status.faultCode');
    AssertEquals_DINT(Expected := 2,
                      Actual := fbNoFeedbackTimeout.status.startCount,
                      Message := 'NoFeedbackTimeout#5 status.startCount');

    // #6, t = 4500 мс — обратная связь пришла: работает
    GVL_S7Clock.tSimNow := T#4500MS;
    fbNoFeedbackTimeout.feedback := TRUE;
    fbNoFeedbackTimeout.reset := FALSE;
    fbNoFeedbackTimeout();
    AssertEquals_BOOL(Expected := TRUE, Actual := fbNoFeedbackTimeout.runCmd, Message := 'NoFeedbackTimeout#6 runCmd');
    AssertEquals_BOOL(Expected := FALSE, Actual := fbNoFeedbackTimeout.fault, Message := 'NoFeedbackTimeout#6 fault');
    AssertEquals_BOOL(Expected := TRUE,
                      Actual := fbNoFeedbackTimeout.status.running,
                      Message := 'NoFeedbackTimeout#6 status.running');
    AssertEquals_BOOL(Expected := FALSE,
                      Actual := fbNoFeedbackTimeout.status.fault,
                      Message := 'NoFeedbackTimeout#6 status.fault');
    AssertEquals_BOOL(Expected := TRUE,
                      Actual := fbNoFeedbackTimeout.status.autoMode,
                      Message := 'NoFeedbackTimeout#6 status.autoMode');
    AssertEquals_INT(Expected := 0,
                     Actual := fbNoFeedbackTimeout.status.faultCode,
                     Message := 'NoFeedbackTimeout#6 status.faultCode');
    AssertEquals_DINT(Expected := 2,
                      Actual := fbNoFeedbackTimeout.status.startCount,
                      Message := 'NoFeedbackTimeout#6 status.startCount');

    // #7, t = 8000 мс — работает
    GVL_S7Clock.tSimNow := T#8000MS;
    fbNoFeedbackTimeout();
    AssertEquals_BOOL(Expected := TRUE, Actual := fbNoFeedbackTimeout.runCmd, Message := 'NoFeedbackTimeout#7 runCmd');
    AssertEquals_BOOL(Expected := FALSE, Actual := fbNoFeedbackTimeout.fault, Message := 'NoFeedbackTimeout#7 fault');
    AssertEquals_BOOL(Expected := TRUE,
                      Actual := fbNoFeedbackTimeout.status.running,
                      Message := 'NoFeedbackTimeout#7 status.running');
    AssertEquals_BOOL(Expected := FALSE,
                      Actual := fbNoFeedbackTimeout.status.fault,
                      Message := 'NoFeedbackTimeout#7 status.fault');
    AssertEquals_BOOL(Expected := TRUE,
                      Actual := fbNoFeedbackTimeout.status.autoMode,
                      Message := 'NoFeedbackTimeout#7 status.autoMode');
    AssertEquals_INT(Expected := 0,
                     Actual := fbNoFeedbackTimeout.status.faultCode,
                     Message := 'NoFeedbackTimeout#7 status.faultCode');
    AssertEquals_DINT(Expected := 2,
                      Actual := fbNoFeedbackTimeout.status.startCount,
                      Message := 'NoFeedbackTimeout#7 status.startCount');

    // #8, t = 8100 мс — стоп
    GVL_S7Clock.tSimNow := T#8100MS;
    fbNoFeedbackTimeout.autoStart := FALSE;
    fbNoFeedbackTimeout();
    AssertEquals_BOOL(Expected := FALSE, Actual := fbNoFeedbackTimeout.runCmd, Message := 'NoFeedbackTimeout#8 runCmd');
    AssertEquals_BOOL(Expected := FALSE, Actual := fbNoFeedbackTimeout.fault, Message := 'NoFeedbackTimeout#8 fault');
    AssertEquals_BOOL(Expected := FALSE,
                      Actual := fbNoFeedbackTimeout.status.running,
                      Message := 'NoFeedbackTimeout#8 status.running');
    AssertEquals_BOOL(Expected := FALSE,
                      Actual := fbNoFeedbackTimeout.status.fault,
                      Message := 'NoFeedbackTimeout#8 status.fault');
    AssertEquals_BOOL(Expected := TRUE,
                      Actual := fbNoFeedbackTimeout.status.autoMode,
                      Message := 'NoFeedbackTimeout#8 status.autoMode');
    AssertEquals_INT(Expected := 0,
                     Actual := fbNoFeedbackTimeout.status.faultCode,
                     Message := 'NoFeedbackTimeout#8 status.faultCode');
    AssertEquals_DINT(Expected := 2,
                      Actual := fbNoFeedbackTimeout.status.startCount,
                      Message := 'NoFeedbackTimeout#8 status.startCount');

    // #9, t = 8300 мс — контактор отпал
    GVL_S7Clock.tSimNow := T#8300MS;
    fbNoFeedbackTimeout.feedback := FALSE;
    fbNoFeedbackTimeout();
    AssertEquals_BOOL(Expected := FALSE, Actual := fbNoFeedbackTimeout.runCmd, Message := 'NoFeedbackTimeout#9 runCmd');
    AssertEquals_BOOL(Expected := FALSE, Actual := fbNoFeedbackTimeout.fault, Message := 'NoFeedbackTimeout#9 fault');
    AssertEquals_BOOL(Expected := FALSE,
                      Actual := fbNoFeedbackTimeout.status.running,
                      Message := 'NoFeedbackTimeout#9 status.running');
    AssertEquals_BOOL(Expected := FALSE,
                      Actual := fbNoFeedbackTimeout.status.fault,
                      Message := 'NoFeedbackTimeout#9 status.fault');
    AssertEquals_BOOL(Expected := TRUE,
                      Actual := fbNoFeedbackTimeout.status.autoMode,
                      Message := 'NoFeedbackTimeout#9 status.autoMode');
    AssertEquals_INT(Expected := 0,
                     Actual := fbNoFeedbackTimeout.status.faultCode,
                     Message := 'NoFeedbackTimeout#9 status.faultCode');
    AssertEquals_DINT(Expected := 2,
                      Actual := fbNoFeedbackTimeout.status.startCount,
                      Message := 'NoFeedbackTimeout#9 status.startCount');

    GVL_S7Clock.xSimulation := FALSE;
END_IF
coUnit.TEST_FINISHED();

(* ---- ThermalTripManual.method.impl.st ---- *)
// AUTO-GENERATED — не редактировать: scenarios/FB_Motor.csv, сценарий ThermalTripManual
coUnit.TEST('ThermalTripManual');
IF NOT xThermalTripManualDone THEN
    xThermalTripManualDone := TRUE;
    GVL_S7Clock.xSimulation := TRUE;

    // #1, t = 0 мс — ручной режим, покой
    GVL_S7Clock.tSimNow := T#0MS;
    fbThermalTripManual.autoMode := FALSE;
    fbThermalTripManual.autoStart := FALSE;
    fbThermalTripManual.manStart := FALSE;
    fbThermalTripManual.manStop := FALSE;
    fbThermalTripManual.feedback := FALSE;
    fbThermalTripManual.thermalOk := TRUE;
    fbThermalTripManual.reset := FALSE;
    fbThermalTripManual.feedbackTime := T#3000MS;
    fbThermalTripManual();
    AssertEquals_BOOL(Expected := FALSE, Actual := fbThermalTripManual.runCmd, Message := 'ThermalTripManual#1 runCmd');
    AssertEquals_BOOL(Expected := FALSE, Actual := fbThermalTripManual.fault, Message := 'ThermalTripManual#1 fault');
    AssertEquals_BOOL(Expected := FALSE,
                      Actual := fbThermalTripManual.status.running,
                      Message := 'ThermalTripManual#1 status.running');
    AssertEquals_BOOL(Expected := FALSE,
                      Actual := fbThermalTripManual.status.fault,
                      Message := 'ThermalTripManual#1 status.fault');
    AssertEquals_BOOL(Expected := FALSE,
                      Actual := fbThermalTripManual.status.autoMode,
                      Message := 'ThermalTripManual#1 status.autoMode');
    AssertEquals_INT(Expected := 0,
                     Actual := fbThermalTripManual.status.faultCode,
                     Message := 'ThermalTripManual#1 status.faultCode');
    AssertEquals_DINT(Expected := 0,
                      Actual := fbThermalTripManual.status.startCount,
                      Message := 'ThermalTripManual#1 status.startCount');

    // #2, t = 100 мс — пуск оператором: пуск №1
    GVL_S7Clock.tSimNow := T#100MS;
    fbThermalTripManual.manStart := TRUE;
    fbThermalTripManual();
    AssertEquals_BOOL(Expected := TRUE, Actual := fbThermalTripManual.runCmd, Message := 'ThermalTripManual#2 runCmd');
    AssertEquals_BOOL(Expected := FALSE, Actual := fbThermalTripManual.fault, Message := 'ThermalTripManual#2 fault');
    AssertEquals_BOOL(Expected := FALSE,
                      Actual := fbThermalTripManual.status.running,
                      Message := 'ThermalTripManual#2 status.running');
    AssertEquals_BOOL(Expected := FALSE,
                      Actual := fbThermalTripManual.status.fault,
                      Message := 'ThermalTripManual#2 status.fault');
    AssertEquals_BOOL(Expected := FALSE,
                      Actual := fbThermalTripManual.status.autoMode,
                      Message := 'ThermalTripManual#2 status.autoMode');
    AssertEquals_INT(Expected := 0,
                     Actual := fbThermalTripManual.status.faultCode,
                     Message := 'ThermalTripManual#2 status.faultCode');
    AssertEquals_DINT(Expected := 1,
                      Actual := fbThermalTripManual.status.startCount,
                      Message := 'ThermalTripManual#2 status.startCount');

    // #3, t = 200 мс — работает
    GVL_S7Clock.tSimNow := T#200MS;
    fbThermalTripManual.manStart := FALSE;
    fbThermalTripManual.feedback := TRUE;
    fbThermalTripManual();
    AssertEquals_BOOL(Expected := TRUE, Actual := fbThermalTripManual.runCmd, Message := 'ThermalTripManual#3 runCmd');
    AssertEquals_BOOL(Expected := FALSE, Actual := fbThermalTripManual.fault, Message := 'ThermalTripManual#3 fault');
    AssertEquals_BOOL(Expected := TRUE,
                      Actual := fbThermalTripManual.status.running,
                      Message := 'ThermalTripManual#3 status.running');
    AssertEquals_BOOL(Expected := FALSE,
                      Actual := fbThermalTripManual.status.fault,
                      Message := 'ThermalTripManual#3 status.fault');
    AssertEquals_BOOL(Expected := FALSE,
                      Actual := fbThermalTripManual.status.autoMode,
                      Message := 'ThermalTripManual#3 status.autoMode');
    AssertEquals_INT(Expected := 0,
                     Actual := fbThermalTripManual.status.faultCode,
                     Message := 'ThermalTripManual#3 status.faultCode');
    AssertEquals_DINT(Expected := 1,
                      Actual := fbThermalTripManual.status.startCount,
                      Message := 'ThermalTripManual#3 status.startCount');

    // #4, t = 1000 мс — тепловая защита: авария 3, ручная защёлка сброшена
    GVL_S7Clock.tSimNow := T#1000MS;
    fbThermalTripManual.thermalOk := FALSE;
    fbThermalTripManual();
    AssertEquals_BOOL(Expected := FALSE, Actual := fbThermalTripManual.runCmd, Message := 'ThermalTripManual#4 runCmd');
    AssertEquals_BOOL(Expected := TRUE, Actual := fbThermalTripManual.fault, Message := 'ThermalTripManual#4 fault');
    AssertEquals_BOOL(Expected := FALSE,
                      Actual := fbThermalTripManual.status.running,
                      Message := 'ThermalTripManual#4 status.running');
    AssertEquals_BOOL(Expected := TRUE,
                      Actual := fbThermalTripManual.status.fault,
                      Message := 'ThermalTripManual#4 status.fault');
    AssertEquals_BOOL(Expected := FALSE,
                      Actual := fbThermalTripManual.status.autoMode,
                      Message := 'ThermalTripManual#4 status.autoMode');
    AssertEquals_INT(Expected := 3,
                     Actual := fbThermalTripManual.status.faultCode,
                     Message := 'ThermalTripManual#4 status.faultCode');
    AssertEquals_DINT(Expected := 1,
                      Actual := fbThermalTripManual.status.startCount,
                      Message := 'ThermalTripManual#4 status.startCount');

    // #5, t = 1500 мс — контактор отпал
    GVL_S7Clock.tSimNow := T#1500MS;
    fbThermalTripManual.feedback := FALSE;
    fbThermalTripManual();
    AssertEquals_BOOL(Expected := FALSE, Actual := fbThermalTripManual.runCmd, Message := 'ThermalTripManual#5 runCmd');
    AssertEquals_BOOL(Expected := TRUE, Actual := fbThermalTripManual.fault, Message := 'ThermalTripManual#5 fault');
    AssertEquals_BOOL(Expected := FALSE,
                      Actual := fbThermalTripManual.status.running,
                      Message := 'ThermalTripManual#5 status.running');
    AssertEquals_BOOL(Expected := TRUE,
                      Actual := fbThermalTripManual.status.fault,
                      Message := 'ThermalTripManual#5 status.fault');
    AssertEquals_BOOL(Expected := FALSE,
                      Actual := fbThermalTripManual.status.autoMode,
                      Message := 'ThermalTripManual#5 status.autoMode');
    AssertEquals_INT(Expected := 3,
                     Actual := fbThermalTripManual.status.faultCode,
                     Message := 'ThermalTripManual#5 status.faultCode');
    AssertEquals_DINT(Expected := 1,
                      Actual := fbThermalTripManual.status.startCount,
                      Message := 'ThermalTripManual#5 status.startCount');

    // #6, t = 2000 мс — сброс при сработавшем реле не действует
    GVL_S7Clock.tSimNow := T#2000MS;
    fbThermalTripManual.reset := TRUE;
    fbThermalTripManual();
    AssertEquals_BOOL(Expected := FALSE, Actual := fbThermalTripManual.runCmd, Message := 'ThermalTripManual#6 runCmd');
    AssertEquals_BOOL(Expected := TRUE, Actual := fbThermalTripManual.fault, Message := 'ThermalTripManual#6 fault');
    AssertEquals_BOOL(Expected := FALSE,
                      Actual := fbThermalTripManual.status.running,
                      Message := 'ThermalTripManual#6 status.running');
    AssertEquals_BOOL(Expected := TRUE,
                      Actual := fbThermalTripManual.status.fault,
                      Message := 'ThermalTripManual#6 status.fault');
    AssertEquals_BOOL(Expected := FALSE,
                      Actual := fbThermalTripManual.status.autoMode,
                      Message := 'ThermalTripManual#6 status.autoMode');
    AssertEquals_INT(Expected := 3,
                     Actual := fbThermalTripManual.status.faultCode,
                     Message := 'ThermalTripManual#6 status.faultCode');
    AssertEquals_DINT(Expected := 1,
                      Actual := fbThermalTripManual.status.startCount,
                      Message := 'ThermalTripManual#6 status.startCount');

    // #7, t = 2500 мс — реле вернулось, авария держится до сброса
    GVL_S7Clock.tSimNow := T#2500MS;
    fbThermalTripManual.thermalOk := TRUE;
    fbThermalTripManual.reset := FALSE;
    fbThermalTripManual();
    AssertEquals_BOOL(Expected := FALSE, Actual := fbThermalTripManual.runCmd, Message := 'ThermalTripManual#7 runCmd');
    AssertEquals_BOOL(Expected := TRUE, Actual := fbThermalTripManual.fault, Message := 'ThermalTripManual#7 fault');
    AssertEquals_BOOL(Expected := FALSE,
                      Actual := fbThermalTripManual.status.running,
                      Message := 'ThermalTripManual#7 status.running');
    AssertEquals_BOOL(Expected := TRUE,
                      Actual := fbThermalTripManual.status.fault,
                      Message := 'ThermalTripManual#7 status.fault');
    AssertEquals_BOOL(Expected := FALSE,
                      Actual := fbThermalTripManual.status.autoMode,
                      Message := 'ThermalTripManual#7 status.autoMode');
    AssertEquals_INT(Expected := 3,
                     Actual := fbThermalTripManual.status.faultCode,
                     Message := 'ThermalTripManual#7 status.faultCode');
    AssertEquals_DINT(Expected := 1,
                      Actual := fbThermalTripManual.status.startCount,
                      Message := 'ThermalTripManual#7 status.startCount');

    // #8, t = 3000 мс — сброс: авария снята, насос не стартует сам
    GVL_S7Clock.tSimNow := T#3000MS;
    fbThermalTripManual.reset := TRUE;
    fbThermalTripManual();
    AssertEquals_BOOL(Expected := FALSE, Actual := fbThermalTripManual.runCmd, Message := 'ThermalTripManual#8 runCmd');
    AssertEquals_BOOL(Expected := FALSE, Actual := fbThermalTripManual.fault, Message := 'ThermalTripManual#8 fault');
    AssertEquals_BOOL(Expected := FALSE,
                      Actual := fbThermalTripManual.status.running,
                      Message := 'ThermalTripManual#8 status.running');
    AssertEquals_BOOL(Expected := FALSE,
                      Actual := fbThermalTripManual.status.fault,
                      Message := 'ThermalTripManual#8 status.fault');
    AssertEquals_BOOL(Expected := FALSE,
                      Actual := fbThermalTripManual.status.autoMode,
                      Message := 'ThermalTripManual#8 status.autoMode');
    AssertEquals_INT(Expected := 0,
                     Actual := fbThermalTripManual.status.faultCode,
                     Message := 'ThermalTripManual#8 status.faultCode');
    AssertEquals_DINT(Expected := 1,
                      Actual := fbThermalTripManual.status.startCount,
                      Message := 'ThermalTripManual#8 status.startCount');

    // #9, t = 3500 мс — новый пуск оператором: пуск №2
    GVL_S7Clock.tSimNow := T#3500MS;
    fbThermalTripManual.manStart := TRUE;
    fbThermalTripManual.reset := FALSE;
    fbThermalTripManual();
    AssertEquals_BOOL(Expected := TRUE, Actual := fbThermalTripManual.runCmd, Message := 'ThermalTripManual#9 runCmd');
    AssertEquals_BOOL(Expected := FALSE, Actual := fbThermalTripManual.fault, Message := 'ThermalTripManual#9 fault');
    AssertEquals_BOOL(Expected := FALSE,
                      Actual := fbThermalTripManual.status.running,
                      Message := 'ThermalTripManual#9 status.running');
    AssertEquals_BOOL(Expected := FALSE,
                      Actual := fbThermalTripManual.status.fault,
                      Message := 'ThermalTripManual#9 status.fault');
    AssertEquals_BOOL(Expected := FALSE,
                      Actual := fbThermalTripManual.status.autoMode,
                      Message := 'ThermalTripManual#9 status.autoMode');
    AssertEquals_INT(Expected := 0,
                     Actual := fbThermalTripManual.status.faultCode,
                     Message := 'ThermalTripManual#9 status.faultCode');
    AssertEquals_DINT(Expected := 2,
                      Actual := fbThermalTripManual.status.startCount,
                      Message := 'ThermalTripManual#9 status.startCount');

    // #10, t = 3600 мс — стоп и пуск одновременно: стоп приоритетнее
    GVL_S7Clock.tSimNow := T#3600MS;
    fbThermalTripManual.manStop := TRUE;
    fbThermalTripManual();
    AssertEquals_BOOL(Expected := FALSE,
                      Actual := fbThermalTripManual.runCmd,
                      Message := 'ThermalTripManual#10 runCmd');
    AssertEquals_BOOL(Expected := FALSE, Actual := fbThermalTripManual.fault, Message := 'ThermalTripManual#10 fault');
    AssertEquals_BOOL(Expected := FALSE,
                      Actual := fbThermalTripManual.status.running,
                      Message := 'ThermalTripManual#10 status.running');
    AssertEquals_BOOL(Expected := FALSE,
                      Actual := fbThermalTripManual.status.fault,
                      Message := 'ThermalTripManual#10 status.fault');
    AssertEquals_BOOL(Expected := FALSE,
                      Actual := fbThermalTripManual.status.autoMode,
                      Message := 'ThermalTripManual#10 status.autoMode');
    AssertEquals_INT(Expected := 0,
                     Actual := fbThermalTripManual.status.faultCode,
                     Message := 'ThermalTripManual#10 status.faultCode');
    AssertEquals_DINT(Expected := 2,
                      Actual := fbThermalTripManual.status.startCount,
                      Message := 'ThermalTripManual#10 status.startCount');

    // #11, t = 3700 мс — покой
    GVL_S7Clock.tSimNow := T#3700MS;
    fbThermalTripManual.manStart := FALSE;
    fbThermalTripManual.manStop := FALSE;
    fbThermalTripManual();
    AssertEquals_BOOL(Expected := FALSE,
                      Actual := fbThermalTripManual.runCmd,
                      Message := 'ThermalTripManual#11 runCmd');
    AssertEquals_BOOL(Expected := FALSE, Actual := fbThermalTripManual.fault, Message := 'ThermalTripManual#11 fault');
    AssertEquals_BOOL(Expected := FALSE,
                      Actual := fbThermalTripManual.status.running,
                      Message := 'ThermalTripManual#11 status.running');
    AssertEquals_BOOL(Expected := FALSE,
                      Actual := fbThermalTripManual.status.fault,
                      Message := 'ThermalTripManual#11 status.fault');
    AssertEquals_BOOL(Expected := FALSE,
                      Actual := fbThermalTripManual.status.autoMode,
                      Message := 'ThermalTripManual#11 status.autoMode');
    AssertEquals_INT(Expected := 0,
                     Actual := fbThermalTripManual.status.faultCode,
                     Message := 'ThermalTripManual#11 status.faultCode');
    AssertEquals_DINT(Expected := 2,
                      Actual := fbThermalTripManual.status.startCount,
                      Message := 'ThermalTripManual#11 status.startCount');

    GVL_S7Clock.xSimulation := FALSE;
END_IF
coUnit.TEST_FINISHED();

(* ---- UnexpectedFeedback.method.impl.st ---- *)
// AUTO-GENERATED — не редактировать: scenarios/FB_Motor.csv, сценарий UnexpectedFeedback
coUnit.TEST('UnexpectedFeedback');
IF NOT xUnexpectedFeedbackDone THEN
    xUnexpectedFeedbackDone := TRUE;
    GVL_S7Clock.xSimulation := TRUE;

    // #1, t = 0 мс — команды нет, обратная связь есть
    GVL_S7Clock.tSimNow := T#0MS;
    fbUnexpectedFeedback.autoMode := TRUE;
    fbUnexpectedFeedback.autoStart := FALSE;
    fbUnexpectedFeedback.manStart := FALSE;
    fbUnexpectedFeedback.manStop := FALSE;
    fbUnexpectedFeedback.feedback := TRUE;
    fbUnexpectedFeedback.thermalOk := TRUE;
    fbUnexpectedFeedback.reset := FALSE;
    fbUnexpectedFeedback.feedbackTime := T#3000MS;
    fbUnexpectedFeedback();
    AssertEquals_BOOL(Expected := FALSE,
                      Actual := fbUnexpectedFeedback.runCmd,
                      Message := 'UnexpectedFeedback#1 runCmd');
    AssertEquals_BOOL(Expected := FALSE, Actual := fbUnexpectedFeedback.fault, Message := 'UnexpectedFeedback#1 fault');
    AssertEquals_BOOL(Expected := FALSE,
                      Actual := fbUnexpectedFeedback.status.running,
                      Message := 'UnexpectedFeedback#1 status.running');
    AssertEquals_BOOL(Expected := FALSE,
                      Actual := fbUnexpectedFeedback.status.fault,
                      Message := 'UnexpectedFeedback#1 status.fault');
    AssertEquals_BOOL(Expected := TRUE,
                      Actual := fbUnexpectedFeedback.status.autoMode,
                      Message := 'UnexpectedFeedback#1 status.autoMode');
    AssertEquals_INT(Expected := 0,
                     Actual := fbUnexpectedFeedback.status.faultCode,
                     Message := 'UnexpectedFeedback#1 status.faultCode');
    AssertEquals_DINT(Expected := 0,
                      Actual := fbUnexpectedFeedback.status.startCount,
                      Message := 'UnexpectedFeedback#1 status.startCount');

    // #2, t = 3200 мс — 3.2 с: авария 4
    GVL_S7Clock.tSimNow := T#3200MS;
    fbUnexpectedFeedback();
    AssertEquals_BOOL(Expected := FALSE,
                      Actual := fbUnexpectedFeedback.runCmd,
                      Message := 'UnexpectedFeedback#2 runCmd');
    AssertEquals_BOOL(Expected := TRUE, Actual := fbUnexpectedFeedback.fault, Message := 'UnexpectedFeedback#2 fault');
    AssertEquals_BOOL(Expected := FALSE,
                      Actual := fbUnexpectedFeedback.status.running,
                      Message := 'UnexpectedFeedback#2 status.running');
    AssertEquals_BOOL(Expected := TRUE,
                      Actual := fbUnexpectedFeedback.status.fault,
                      Message := 'UnexpectedFeedback#2 status.fault');
    AssertEquals_BOOL(Expected := TRUE,
                      Actual := fbUnexpectedFeedback.status.autoMode,
                      Message := 'UnexpectedFeedback#2 status.autoMode');
    AssertEquals_INT(Expected := 4,
                     Actual := fbUnexpectedFeedback.status.faultCode,
                     Message := 'UnexpectedFeedback#2 status.faultCode');
    AssertEquals_DINT(Expected := 0,
                      Actual := fbUnexpectedFeedback.status.startCount,
                      Message := 'UnexpectedFeedback#2 status.startCount');

    // #3, t = 4000 мс — сброс: таймер всё ещё в Q — авария 4 снова в том же вызове
    GVL_S7Clock.tSimNow := T#4000MS;
    fbUnexpectedFeedback.reset := TRUE;
    fbUnexpectedFeedback();
    AssertEquals_BOOL(Expected := FALSE,
                      Actual := fbUnexpectedFeedback.runCmd,
                      Message := 'UnexpectedFeedback#3 runCmd');
    AssertEquals_BOOL(Expected := TRUE, Actual := fbUnexpectedFeedback.fault, Message := 'UnexpectedFeedback#3 fault');
    AssertEquals_BOOL(Expected := FALSE,
                      Actual := fbUnexpectedFeedback.status.running,
                      Message := 'UnexpectedFeedback#3 status.running');
    AssertEquals_BOOL(Expected := TRUE,
                      Actual := fbUnexpectedFeedback.status.fault,
                      Message := 'UnexpectedFeedback#3 status.fault');
    AssertEquals_BOOL(Expected := TRUE,
                      Actual := fbUnexpectedFeedback.status.autoMode,
                      Message := 'UnexpectedFeedback#3 status.autoMode');
    AssertEquals_INT(Expected := 4,
                     Actual := fbUnexpectedFeedback.status.faultCode,
                     Message := 'UnexpectedFeedback#3 status.faultCode');
    AssertEquals_DINT(Expected := 0,
                      Actual := fbUnexpectedFeedback.status.startCount,
                      Message := 'UnexpectedFeedback#3 status.startCount');

    // #4, t = 4500 мс — контактор отпал, авария держится
    GVL_S7Clock.tSimNow := T#4500MS;
    fbUnexpectedFeedback.feedback := FALSE;
    fbUnexpectedFeedback.reset := FALSE;
    fbUnexpectedFeedback();
    AssertEquals_BOOL(Expected := FALSE,
                      Actual := fbUnexpectedFeedback.runCmd,
                      Message := 'UnexpectedFeedback#4 runCmd');
    AssertEquals_BOOL(Expected := TRUE, Actual := fbUnexpectedFeedback.fault, Message := 'UnexpectedFeedback#4 fault');
    AssertEquals_BOOL(Expected := FALSE,
                      Actual := fbUnexpectedFeedback.status.running,
                      Message := 'UnexpectedFeedback#4 status.running');
    AssertEquals_BOOL(Expected := TRUE,
                      Actual := fbUnexpectedFeedback.status.fault,
                      Message := 'UnexpectedFeedback#4 status.fault');
    AssertEquals_BOOL(Expected := TRUE,
                      Actual := fbUnexpectedFeedback.status.autoMode,
                      Message := 'UnexpectedFeedback#4 status.autoMode');
    AssertEquals_INT(Expected := 4,
                     Actual := fbUnexpectedFeedback.status.faultCode,
                     Message := 'UnexpectedFeedback#4 status.faultCode');
    AssertEquals_DINT(Expected := 0,
                      Actual := fbUnexpectedFeedback.status.startCount,
                      Message := 'UnexpectedFeedback#4 status.startCount');

    // #5, t = 5000 мс — сброс: авария снята
    GVL_S7Clock.tSimNow := T#5000MS;
    fbUnexpectedFeedback.reset := TRUE;
    fbUnexpectedFeedback();
    AssertEquals_BOOL(Expected := FALSE,
                      Actual := fbUnexpectedFeedback.runCmd,
                      Message := 'UnexpectedFeedback#5 runCmd');
    AssertEquals_BOOL(Expected := FALSE, Actual := fbUnexpectedFeedback.fault, Message := 'UnexpectedFeedback#5 fault');
    AssertEquals_BOOL(Expected := FALSE,
                      Actual := fbUnexpectedFeedback.status.running,
                      Message := 'UnexpectedFeedback#5 status.running');
    AssertEquals_BOOL(Expected := FALSE,
                      Actual := fbUnexpectedFeedback.status.fault,
                      Message := 'UnexpectedFeedback#5 status.fault');
    AssertEquals_BOOL(Expected := TRUE,
                      Actual := fbUnexpectedFeedback.status.autoMode,
                      Message := 'UnexpectedFeedback#5 status.autoMode');
    AssertEquals_INT(Expected := 0,
                     Actual := fbUnexpectedFeedback.status.faultCode,
                     Message := 'UnexpectedFeedback#5 status.faultCode');
    AssertEquals_DINT(Expected := 0,
                      Actual := fbUnexpectedFeedback.status.startCount,
                      Message := 'UnexpectedFeedback#5 status.startCount');

    // #6, t = 5500 мс — пуск №1
    GVL_S7Clock.tSimNow := T#5500MS;
    fbUnexpectedFeedback.autoStart := TRUE;
    fbUnexpectedFeedback.reset := FALSE;
    fbUnexpectedFeedback();
    AssertEquals_BOOL(Expected := TRUE,
                      Actual := fbUnexpectedFeedback.runCmd,
                      Message := 'UnexpectedFeedback#6 runCmd');
    AssertEquals_BOOL(Expected := FALSE, Actual := fbUnexpectedFeedback.fault, Message := 'UnexpectedFeedback#6 fault');
    AssertEquals_BOOL(Expected := FALSE,
                      Actual := fbUnexpectedFeedback.status.running,
                      Message := 'UnexpectedFeedback#6 status.running');
    AssertEquals_BOOL(Expected := FALSE,
                      Actual := fbUnexpectedFeedback.status.fault,
                      Message := 'UnexpectedFeedback#6 status.fault');
    AssertEquals_BOOL(Expected := TRUE,
                      Actual := fbUnexpectedFeedback.status.autoMode,
                      Message := 'UnexpectedFeedback#6 status.autoMode');
    AssertEquals_INT(Expected := 0,
                     Actual := fbUnexpectedFeedback.status.faultCode,
                     Message := 'UnexpectedFeedback#6 status.faultCode');
    AssertEquals_DINT(Expected := 1,
                      Actual := fbUnexpectedFeedback.status.startCount,
                      Message := 'UnexpectedFeedback#6 status.startCount');

    // #7, t = 6000 мс — работает
    GVL_S7Clock.tSimNow := T#6000MS;
    fbUnexpectedFeedback.feedback := TRUE;
    fbUnexpectedFeedback();
    AssertEquals_BOOL(Expected := TRUE,
                      Actual := fbUnexpectedFeedback.runCmd,
                      Message := 'UnexpectedFeedback#7 runCmd');
    AssertEquals_BOOL(Expected := FALSE, Actual := fbUnexpectedFeedback.fault, Message := 'UnexpectedFeedback#7 fault');
    AssertEquals_BOOL(Expected := TRUE,
                      Actual := fbUnexpectedFeedback.status.running,
                      Message := 'UnexpectedFeedback#7 status.running');
    AssertEquals_BOOL(Expected := FALSE,
                      Actual := fbUnexpectedFeedback.status.fault,
                      Message := 'UnexpectedFeedback#7 status.fault');
    AssertEquals_BOOL(Expected := TRUE,
                      Actual := fbUnexpectedFeedback.status.autoMode,
                      Message := 'UnexpectedFeedback#7 status.autoMode');
    AssertEquals_INT(Expected := 0,
                     Actual := fbUnexpectedFeedback.status.faultCode,
                     Message := 'UnexpectedFeedback#7 status.faultCode');
    AssertEquals_DINT(Expected := 1,
                      Actual := fbUnexpectedFeedback.status.startCount,
                      Message := 'UnexpectedFeedback#7 status.startCount');

    GVL_S7Clock.xSimulation := FALSE;
END_IF
coUnit.TEST_FINISHED();
